// TIA Portal project "FactoryIO_Template_S7-1200_V15_V18_5" (V18)
// Vorlageprojekt für das Buch mit Zielsystem S7-1200

(* hardware
DEVICE "S7-1200-Station_1"  S7-1200 Station
   slot 0: "Baugruppenträger_0"  Rack  V1.0
   slot 1: "PLC_1"  CPU 1214C AC/DC/Rly  6ES7 214-1BG40-0XB0  V4.6
   slot 2: "AQ 4x14BIT_1"  6ES7 232-4HD32-0XB0  V2.1
*)

// ===== PLC "PLC_1"  CPU 1214C AC/DC/Rly =====

VAR_GLOBAL   // PLC tag table "Standard-Variablentabelle"
   "Start_Butonu" AT %I0.0 : Bool;
   "Stop_Butonu" AT %I0.1 : Bool;
   "Reset_Butonu" AT %I0.2 : Bool;
   "Doldurma_Miktarı" AT %IW30 : Int;
   "Seviye_Tespit_Sensörü" AT %IW32 : Int;
   "Start_Lambası" AT %Q0.0 : Bool;
   "Stop_Lambası" AT %Q0.1 : Bool;
   "Reset_Lambası" AT %Q0.2 : Bool;
   "Doldurma_Valfi" AT %QW30 : Int;
   "Boşaltma_Valfi" AT %QW32 : Int;
   "Hedef_Seviye" AT %QW34 : Int;
   "Gerçek_Seviye" AT %QW36 : Int;
   "Sistem Genel Start" AT %M10.0 : Bool;
   "Tag_1" AT %MW20 : Int;
   "Tag_2" AT %MD22 : Real;
   "Sıvı_Seviyesi" AT %MD26 : Real;
   "Tag_4" AT %MW12 : Int;
END_VAR

// folder: System blocks/Program resources

DATA_BLOCK "Timer-1"   // DB1
{ S7_Optimized_Access := 'TRUE' }
AUTHOR : Simatic
FAMILY : IEC
NAME : IEC_TMR
VERSION : 1.0
// stored: InstanceOfName IEC_TIMER
"IEC_TIMER"
BEGIN
END_DATA_BLOCK

// folder: (top level)

FUNCTION "MHJ-PLC-Lab-Function-S71200" : Void   // FC9000, SCL
{ S7_Optimized_Access := 'TRUE' }
VERSION : 0.1
   VAR_TEMP
      rdTimeReturn : Int;
      outputTime : DTL;
      SyncVal : Byte;
      forVal : Int;
      forVal_2 : Int;
      Value : Byte;
   END_VAR
   VAR CONSTANT
      CompVal : Byte := 16#34;
      Value_01 : Byte := 16#11;
      Value_01_DW : DWord := 16#A165_D992;
      Value_02_DW : DWord := 16#58BE_4401;
   END_VAR
BEGIN

   #Value:=PEEK(area := 16#82,
        dbNumber := 0,
        byteOffset := 511);
   #Value := #Value + 1;

   POKE(area := 16#82,
        dbNumber := 0,
        byteOffset := 511,
        value := #Value);

   POKE(area:=16#81,
        dbNumber:=0,
        byteOffset:=1016,
        value:=#Value_01_DW);
   POKE(area := 16#81,
        dbNumber := 0,
        byteOffset := 1020,
        value := #Value_02_DW);

   POKE(area := 16#81,
        dbNumber := 0,
        byteOffset := 511,
        value := B#16#00);

   FOR #forVal := 0 TO 120 DO
       FOR #forVal_2:=0 TO 10 DO
           #rdTimeReturn:=RD_SYS_T(#outputTime);
           #rdTimeReturn := WR_SYS_T(#outputTime);
           #rdTimeReturn := RD_SYS_T(#outputTime);
           #rdTimeReturn := WR_SYS_T(#outputTime);
       END_FOR;
       #SyncVal:= PEEK(area := 16#81,
                      dbNumber := 0,
                      byteOffset := 511);
       IF #SyncVal = #CompVal THEN
          GOTO M_1;
       END_IF;
   END_FOR;
   RETURN;

   M_1:
   POKE(area := 16#81,
        dbNumber := 0,
        byteOffset := 511,
        value := B#16#0);
END_FUNCTION

ORGANIZATION_BLOCK "Main"   // OB1, LAD, ProgramCycle
TITLE = "Main Program Sweep (Cycle)"
{ S7_Optimized_Access := 'TRUE' }
VERSION : 0.1
   VAR_INPUT
      Initial_Call : Bool;   // Initial call of this OB
      Remanence : Bool;   // =True, if remanent data are available
   END_VAR
BEGIN

REGION Network 1: Konnektierungsbaustein für PLC-Lab / FACTORY I/O HABERLEŞME BAĞLANTISI
   // Im Netzwerk 1 wird der Konnektierungsbaustein für PLC-Lab aufgerufen.
   // Dieser Aufruf darf nicht entfernt werden!
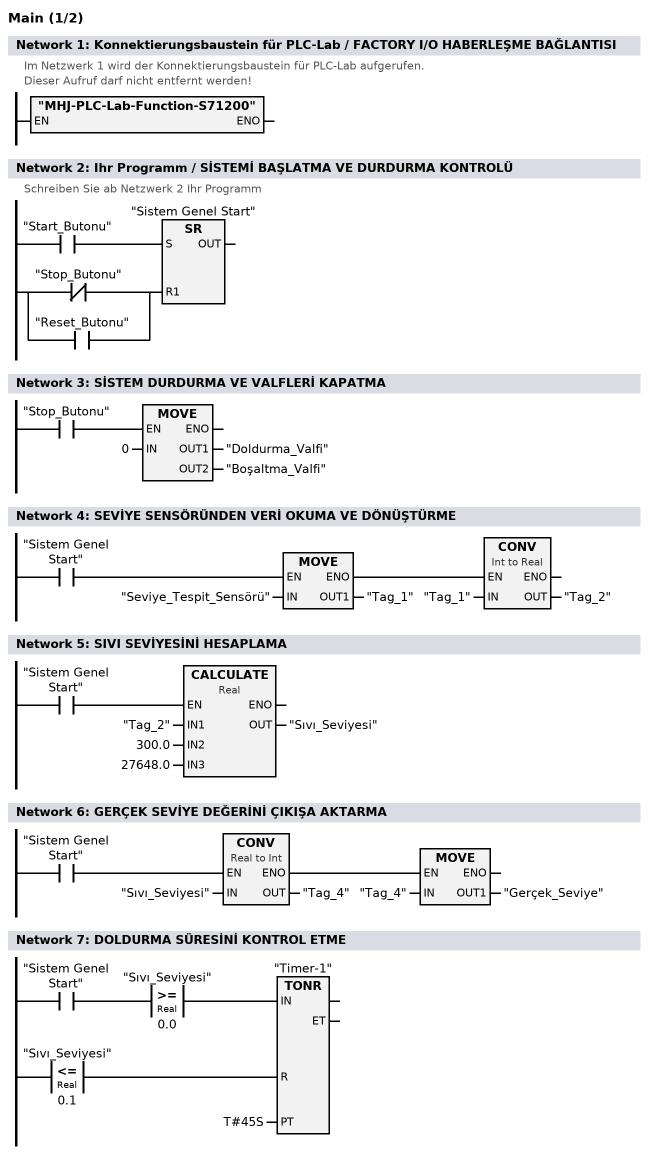
   RUNG wire#powerrail
      "MHJ-PLC-Lab-Function-S71200"()
   END_RUNG
   // the same network as SCL:
   "MHJ-PLC-Lab-Function-S71200"();
END_REGION

REGION Network 2: Ihr Programm / SİSTEMİ BAŞLATMA VE DURDURMA KONTROLÜ
   // Schreiben Sie ab Netzwerk 2 Ihr Programm
   RUNG wire#powerrail
      Contact( "Start_Butonu" )
      S_SR(operand := "Sistem Genel Start", r1 := wire#w1)
   END_RUNG
   RUNG wire#powerrail
      I_Contact( "Stop_Butonu" )
   END_RUNG wire#w1
   RUNG wire#powerrail
      Contact( "Reset_Butonu" )
   END_RUNG wire#w1
   // the same network as SCL:
   IF "Start_Butonu" THEN
       "Sistem Genel Start" := TRUE;   // SR flip-flop
   END_IF;
   IF NOT "Stop_Butonu" OR "Reset_Butonu" THEN "Sistem Genel Start" := FALSE; END_IF;
END_REGION

REGION Network 3: SİSTEM DURDURMA VE VALFLERİ KAPATMA
   RUNG wire#powerrail
      Contact( "Stop_Butonu" )
      Move(in := 0, out1 => "Doldurma_Valfi", out2 => "Boşaltma_Valfi")
   END_RUNG
   // the same network as SCL:
   IF "Stop_Butonu" THEN
       "Doldurma_Valfi" := 0;
       "Boşaltma_Valfi" := 0;
   END_IF;
END_REGION

REGION Network 4: SEVİYE SENSÖRÜNDEN VERİ OKUMA VE DÖNÜŞTÜRME
   RUNG wire#powerrail
      Contact( "Sistem Genel Start" )
      Move(in := "Seviye_Tespit_Sensörü", out1 => "Tag_1")
      { S7_Templates := "[SrcType := Int, DestType := Real]" } Convert(in := "Tag_1", out => "Tag_2")
   END_RUNG
   // the same network as SCL:
   IF "Sistem Genel Start" THEN
       "Tag_1" := "Seviye_Tespit_Sensörü";
       "Tag_2" := INT_TO_REAL("Tag_1");
   END_IF;
END_REGION

REGION Network 5: SIVI SEVİYESİNİ HESAPLAMA
   RUNG wire#powerrail
      Contact( "Sistem Genel Start" )
      { S7_Templates := "SrcType := Real"; S7_Expression := "(IN1*IN2)/IN3" } Calculate(in1 := "Tag_2", in2 := 300.0, in3 := 27648.0, out => "Sıvı_Seviyesi")
   END_RUNG
   // the same network as SCL:
   IF "Sistem Genel Start" THEN "Sıvı_Seviyesi" := ("Tag_2"*300.0)/27648.0; END_IF;
END_REGION

REGION Network 6: GERÇEK SEVİYE DEĞERİNİ ÇIKIŞA AKTARMA
   RUNG wire#powerrail
      Contact( "Sistem Genel Start" )
      { S7_Templates := "[SrcType := Real, DestType := Int]" } Convert(in := "Sıvı_Seviyesi", out => "Tag_4")
      Move(in := "Tag_4", out1 => "Gerçek_Seviye")
   END_RUNG
   // the same network as SCL:
   IF "Sistem Genel Start" THEN
       "Tag_4" := REAL_TO_INT("Sıvı_Seviyesi");
       "Gerçek_Seviye" := "Tag_4";
   END_IF;
END_REGION

REGION Network 7: DOLDURMA SÜRESİNİ KONTROL ETME
   "Timer-1".TONR(IN := "Sistem Genel Start" AND ("Sıvı_Seviyesi" >= 0.0),
                  R := "Sıvı_Seviyesi" <= 0.1,
                  PT := T#45S);
END_REGION

REGION Network 8: TANK DOLDURMA KONTROLÜ
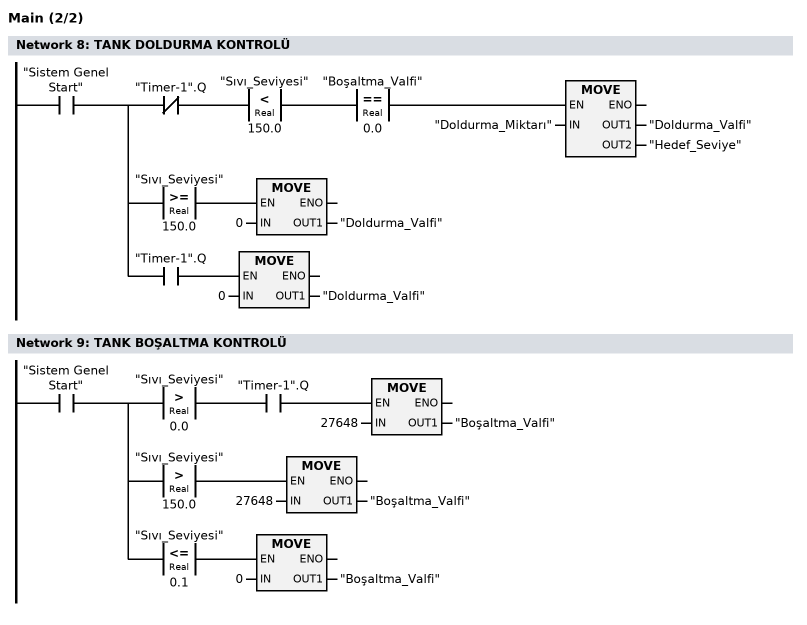
   RUNG wire#powerrail
      Contact( "Sistem Genel Start" )
      wire#w1
      I_Contact( "Timer-1".Q )
      { S7_Templates := "SrcType := Real" } LT_Contact(in1 := "Sıvı_Seviyesi", in2 := 150.0)
      { S7_Templates := "SrcType := Real" } EQ_Contact(in1 := "Boşaltma_Valfi", in2 := 0.0)
      Move(in := "Doldurma_Miktarı", out1 => "Doldurma_Valfi", out2 => "Hedef_Seviye")
   END_RUNG
   RUNG wire#w1
      { S7_Templates := "SrcType := Real" } GE_Contact(in1 := "Sıvı_Seviyesi", in2 := 150.0)
      Move(in := 0, out1 => "Doldurma_Valfi")
   END_RUNG
   RUNG wire#w1
      Contact( "Timer-1".Q )
      Move(in := 0, out1 => "Doldurma_Valfi")
   END_RUNG
   // the same network as SCL:
   IF "Sistem Genel Start" AND NOT "Timer-1".Q AND ("Sıvı_Seviyesi" < 150.0) AND ("Boşaltma_Valfi" = 0.0) THEN
       "Doldurma_Valfi" := "Doldurma_Miktarı";
       "Hedef_Seviye" := "Doldurma_Miktarı";
   END_IF;
   IF "Sistem Genel Start" AND ("Sıvı_Seviyesi" >= 150.0) THEN "Doldurma_Valfi" := 0; END_IF;
   IF "Sistem Genel Start" AND "Timer-1".Q THEN "Doldurma_Valfi" := 0; END_IF;
END_REGION

REGION Network 9: TANK BOŞALTMA KONTROLÜ
   RUNG wire#powerrail
      Contact( "Sistem Genel Start" )
      wire#w1
      { S7_Templates := "SrcType := Real" } GT_Contact(in1 := "Sıvı_Seviyesi", in2 := 0.0)
      Contact( "Timer-1".Q )
      Move(in := 27648, out1 => "Boşaltma_Valfi")
   END_RUNG
   RUNG wire#w1
      { S7_Templates := "SrcType := Real" } GT_Contact(in1 := "Sıvı_Seviyesi", in2 := 150.0)
      Move(in := 27648, out1 => "Boşaltma_Valfi")
   END_RUNG
   RUNG wire#w1
      { S7_Templates := "SrcType := Real" } LE_Contact(in1 := "Sıvı_Seviyesi", in2 := 0.1)
      Move(in := 0, out1 => "Boşaltma_Valfi")
   END_RUNG
   // the same network as SCL:
   IF "Sistem Genel Start" AND ("Sıvı_Seviyesi" > 0.0) AND "Timer-1".Q THEN
       "Boşaltma_Valfi" := 27648;
   END_IF;
   IF "Sistem Genel Start" AND ("Sıvı_Seviyesi" > 150.0) THEN "Boşaltma_Valfi" := 27648; END_IF;
   IF "Sistem Genel Start" AND ("Sıvı_Seviyesi" <= 0.1) THEN "Boşaltma_Valfi" := 0; END_IF;
END_REGION
END_ORGANIZATION_BLOCK